FUNCTION_BLOCK "OP5_Pressure_Interlocks"
{ S7_Optimized_Access := 'TRUE' }
VERSION : 0.1
   VAR
      State {InstructionName := 'Program_Alarm'; LibVersion := '1.0'} : Program_Alarm;
      PRECOND_01 : Bool;
      PRECOND_02 : Bool;
      PRECOND_03 : Bool;
      PRECOND_04 : Bool;
      PRECOND_05 : Bool;
      PRECOND_06 : Bool;
      PRECOND_07 : Bool;
      PRECOND_08 : Bool;
      PRECOND_09 : Bool;
      PRECOND_10 : Bool;
      PRECOND_11 : Bool;
      PRECOND_12 : Bool;
      PRECOND_13 : Bool;
      PRECOND_14 : Bool;
      PRECOND_15 : Bool;
      PRECOND_16 : Bool;
      PRECOND_17 : Bool;
      PRECOND_18 : Bool;
      PRECOND_19 : Bool;
      PRECOND_20 : Bool;
      PRECOND_21 : Bool;
      PRECOND_22 : Bool;
      PRECOND_23 : Bool;
      PRECOND_24 : Bool;
      PRECOND_25 : Bool;
      PRECOND_26 : Bool;
      PRECOND_27 : Bool;
      PRECOND_28 : Bool;
      PRECOND_29 : Bool;
      PRECOND_30 : Bool;
      PRECOND_31 : Bool;
      PRECOND_32 : Bool;
      PRECOND_33 : Bool;
      PRECOND_34 : Bool;
      PRECOND_35 : Bool;
      PRECOND_36 : Bool;
      PRECOND_37 : Bool;
      PRECOND_38 : Bool;
      PRECOND_39 : Bool;
      PRECOND_40 : Bool;
      PRECOND_41 : Bool;
      PRECOND_42 : Bool;
      PRECOND_43 : Bool;
      PRECOND_44 : Bool;
      PRECOND_45 : Bool;
      PRECOND_46 : Bool;
      PRECOND_47 : Bool;
      PRECOND_48 : Bool;
      PRECOND_49 : Bool;
      PRECOND_50 : Bool;
      PH_Vent_PRECOND_01 : Bool;
      PH_Vent_PRECOND_02 : Bool;
      PH_Vent_PRECOND_03 : Bool;
      PH_Vent_PRECOND_04 : Bool;
      PH_Vent_PRECOND_05 : Bool;
      PH_Vent_PRECOND_06 : Bool;
      PH_Vent_PRECOND_07 : Bool;
      PH_Vent_PRECOND_08 : Bool;
      PH_Vent_PRECOND_09 : Bool;
      PH_Vent_PRECOND_10 : Bool;
      PH_Vent_PRECOND_11 : Bool;
      PH_Vent_PRECOND_12 : Bool;
      PH_Vent_PRECOND_13 : Bool;
      PH_Vent_PRECOND_14 : Bool;
      PH_Vent_PRECOND_15 : Bool;
      PH_Vent_PRECOND_16 : Bool;
      PH_Vent_PRECOND_17 : Bool;
      PH_Vent_PRECOND_18 : Bool;
      PH_Vent_PRECOND_19 : Bool;
      PH_Vent_PRECOND_20 : Bool;
      PH_Vent_PRECOND_21 : Bool;
      PH_Vent_PRECOND_22 : Bool;
      PH_Vent_PRECOND_23 : Bool;
      PH_Vent_PRECOND_24 : Bool;
      PH_Vent_PRECOND_25 : Bool;
      PH_Vent_PRECOND_26 : Bool;
      PH_Vent_PRECOND_27 : Bool;
      PH_Vent_PRECOND_28 : Bool;
      PH_Vent_PRECOND_29 : Bool;
      PH_Vent_PRECOND_30 : Bool;
      PH_Vent_PRECOND_31 : Bool;
      PH_Vent_PRECOND_32 : Bool;
      PH_Vent_PRECOND_33 : Bool;
      PH_Vent_PRECOND_34 : Bool;
      PH_Vent_PRECOND_35 : Bool;
      PH_Vent_PRECOND_36 : Bool;
      PH_Vent_PRECOND_37 : Bool;
      PH_Vent_PRECOND_38 : Bool;
      PH_Vent_PRECOND_39 : Bool;
      PH_Vent_PRECOND_40 : Bool;
      PH_Vent_PRECOND_41 : Bool;
      PH_Vent_PRECOND_42 : Bool;
      PH_Vent_PRECOND_43 : Bool;
      PH_Vent_PRECOND_44 : Bool;
      PH_Vent_PRECOND_45 : Bool;
      PH_Vent_PRECOND_46 : Bool;
      PH_Vent_PRECOND_47 : Bool;
      PH_Vent_PRECOND_48 : Bool;
      PH_Vent_PRECOND_49 : Bool;
      PH_Vent_PRECOND_50 : Bool;
      PH_Fill_PRECOND_01 : Bool;
      PH_Fill_PRECOND_02 : Bool;
      PH_Fill_PRECOND_03 : Bool;
      PH_Fill_PRECOND_04 : Bool;
      PH_Fill_PRECOND_05 : Bool;
      PH_Fill_PRECOND_06 : Bool;
      PH_Fill_PRECOND_07 : Bool;
      PH_Fill_PRECOND_08 : Bool;
      PH_Fill_PRECOND_09 : Bool;
      PH_Fill_PRECOND_10 : Bool;
      PH_Fill_PRECOND_11 : Bool;
      PH_Fill_PRECOND_12 : Bool;
      PH_Fill_PRECOND_13 : Bool;
      PH_Fill_PRECOND_14 : Bool;
      PH_Fill_PRECOND_15 : Bool;
      PH_Fill_PRECOND_16 : Bool;
      PH_Fill_PRECOND_17 : Bool;
      PH_Fill_PRECOND_18 : Bool;
      PH_Fill_PRECOND_19 : Bool;
      PH_Fill_PRECOND_20 : Bool;
      PH_Fill_PRECOND_21 : Bool;
      PH_Fill_PRECOND_22 : Bool;
      PH_Fill_PRECOND_23 : Bool;
      PH_Fill_PRECOND_24 : Bool;
      PH_Fill_PRECOND_25 : Bool;
      PH_Fill_PRECOND_26 : Bool;
      PH_Fill_PRECOND_27 : Bool;
      PH_Fill_PRECOND_28 : Bool;
      PH_Fill_PRECOND_29 : Bool;
      PH_Fill_PRECOND_30 : Bool;
      PH_Fill_PRECOND_31 : Bool;
      PH_Fill_PRECOND_32 : Bool;
      PH_Fill_PRECOND_33 : Bool;
      PH_Fill_PRECOND_34 : Bool;
      PH_Fill_PRECOND_35 : Bool;
      PH_Fill_PRECOND_36 : Bool;
      PH_Fill_PRECOND_37 : Bool;
      PH_Fill_PRECOND_38 : Bool;
      PH_Fill_PRECOND_39 : Bool;
      PH_Fill_PRECOND_40 : Bool;
      PH_Fill_PRECOND_41 : Bool;
      PH_Fill_PRECOND_42 : Bool;
      PH_Fill_PRECOND_43 : Bool;
      PH_Fill_PRECOND_44 : Bool;
      PH_Fill_PRECOND_45 : Bool;
      PH_Fill_PRECOND_46 : Bool;
      PH_Fill_PRECOND_47 : Bool;
      PH_Fill_PRECOND_48 : Bool;
      PH_Fill_PRECOND_49 : Bool;
      PH_Fill_PRECOND_50 : Bool;
   END_VAR

BEGIN
   REGION Function
      // here all interlocks for this operation will be defined
      // Later FALSE assignments execute every scan. Adjust them when adding calculated interlocks.
   END_REGION

   REGION General Interlocks
      #PRECOND_01 := FALSE;
      #PRECOND_02 := FALSE;
      #PRECOND_03 := FALSE;
      #PRECOND_04 := FALSE;
      #PRECOND_05 := FALSE;
      #PRECOND_06 := FALSE;
      #PRECOND_07 := FALSE;
      #PRECOND_08 := FALSE;
      #PRECOND_09 := FALSE;
      #PRECOND_10 := FALSE;
      #PRECOND_11 := FALSE;
      #PRECOND_12 := FALSE;
      #PRECOND_13 := FALSE;
      #PRECOND_14 := FALSE;
      #PRECOND_15 := FALSE;
      #PRECOND_16 := FALSE;
      #PRECOND_17 := FALSE;
      #PRECOND_18 := FALSE;
      #PRECOND_19 := FALSE;
      #PRECOND_20 := FALSE;
      #PRECOND_21 := FALSE;
      #PRECOND_22 := FALSE;
      #PRECOND_23 := FALSE;
      #PRECOND_24 := FALSE;
      #PRECOND_25 := FALSE;
      #PRECOND_26 := FALSE;
      #PRECOND_27 := FALSE;
      #PRECOND_28 := FALSE;
      #PRECOND_29 := FALSE;
      #PRECOND_30 := FALSE;
      #PRECOND_31 := FALSE;
      #PRECOND_32 := FALSE;
      #PRECOND_33 := FALSE;
      #PRECOND_34 := FALSE;
      #PRECOND_35 := FALSE;
      #PRECOND_36 := FALSE;
      #PRECOND_37 := FALSE;
      #PRECOND_38 := FALSE;
      #PRECOND_39 := FALSE;
      #PRECOND_40 := FALSE;
      #PRECOND_41 := FALSE;
      #PRECOND_42 := FALSE;
      #PRECOND_43 := FALSE;
      #PRECOND_44 := FALSE;
      #PRECOND_45 := FALSE;
      #PRECOND_46 := FALSE;
      #PRECOND_47 := FALSE;
      #PRECOND_48 := FALSE;
      #PRECOND_49 := FALSE;
      #PRECOND_50 := FALSE;
   END_REGION

   REGION PH_Vent Interlocks
      #PH_Vent_PRECOND_01 := FALSE;
      #PH_Vent_PRECOND_02 := FALSE;
      #PH_Vent_PRECOND_03 := FALSE;
      #PH_Vent_PRECOND_04 := FALSE;
      #PH_Vent_PRECOND_05 := FALSE;
      #PH_Vent_PRECOND_06 := FALSE;
      #PH_Vent_PRECOND_07 := FALSE;
      #PH_Vent_PRECOND_08 := FALSE;
      #PH_Vent_PRECOND_09 := FALSE;
      #PH_Vent_PRECOND_10 := FALSE;
      #PH_Vent_PRECOND_11 := FALSE;
      #PH_Vent_PRECOND_12 := FALSE;
      #PH_Vent_PRECOND_13 := FALSE;
      #PH_Vent_PRECOND_14 := FALSE;
      #PH_Vent_PRECOND_15 := FALSE;
      #PH_Vent_PRECOND_16 := FALSE;
      #PH_Vent_PRECOND_17 := FALSE;
      #PH_Vent_PRECOND_18 := FALSE;
      #PH_Vent_PRECOND_19 := FALSE;
      #PH_Vent_PRECOND_20 := FALSE;
      #PH_Vent_PRECOND_21 := FALSE;
      #PH_Vent_PRECOND_22 := FALSE;
      #PH_Vent_PRECOND_23 := FALSE;
      #PH_Vent_PRECOND_24 := FALSE;
      #PH_Vent_PRECOND_25 := FALSE;
      #PH_Vent_PRECOND_26 := FALSE;
      #PH_Vent_PRECOND_27 := FALSE;
      #PH_Vent_PRECOND_28 := FALSE;
      #PH_Vent_PRECOND_29 := FALSE;
      #PH_Vent_PRECOND_30 := FALSE;
      #PH_Vent_PRECOND_31 := FALSE;
      #PH_Vent_PRECOND_32 := FALSE;
      #PH_Vent_PRECOND_33 := FALSE;
      #PH_Vent_PRECOND_34 := FALSE;
      #PH_Vent_PRECOND_35 := FALSE;
      #PH_Vent_PRECOND_36 := FALSE;
      #PH_Vent_PRECOND_37 := FALSE;
      #PH_Vent_PRECOND_38 := FALSE;
      #PH_Vent_PRECOND_39 := FALSE;
      #PH_Vent_PRECOND_40 := FALSE;
      #PH_Vent_PRECOND_41 := FALSE;
      #PH_Vent_PRECOND_42 := FALSE;
      #PH_Vent_PRECOND_43 := FALSE;
      #PH_Vent_PRECOND_44 := FALSE;
      #PH_Vent_PRECOND_45 := FALSE;
      #PH_Vent_PRECOND_46 := FALSE;
      #PH_Vent_PRECOND_47 := FALSE;
      #PH_Vent_PRECOND_48 := FALSE;
      #PH_Vent_PRECOND_49 := FALSE;
      #PH_Vent_PRECOND_50 := FALSE;
   END_REGION

   REGION PH_Fill Interlocks
      #PH_Fill_PRECOND_01 := FALSE;
      #PH_Fill_PRECOND_02 := FALSE;
      #PH_Fill_PRECOND_03 := FALSE;
      #PH_Fill_PRECOND_04 := FALSE;
      #PH_Fill_PRECOND_05 := FALSE;
      #PH_Fill_PRECOND_06 := FALSE;
      #PH_Fill_PRECOND_07 := FALSE;
      #PH_Fill_PRECOND_08 := FALSE;
      #PH_Fill_PRECOND_09 := FALSE;
      #PH_Fill_PRECOND_10 := FALSE;
      #PH_Fill_PRECOND_11 := FALSE;
      #PH_Fill_PRECOND_12 := FALSE;
      #PH_Fill_PRECOND_13 := FALSE;
      #PH_Fill_PRECOND_14 := FALSE;
      #PH_Fill_PRECOND_15 := FALSE;
      #PH_Fill_PRECOND_16 := FALSE;
      #PH_Fill_PRECOND_17 := FALSE;
      #PH_Fill_PRECOND_18 := FALSE;
      #PH_Fill_PRECOND_19 := FALSE;
      #PH_Fill_PRECOND_20 := FALSE;
      #PH_Fill_PRECOND_21 := FALSE;
      #PH_Fill_PRECOND_22 := FALSE;
      #PH_Fill_PRECOND_23 := FALSE;
      #PH_Fill_PRECOND_24 := FALSE;
      #PH_Fill_PRECOND_25 := FALSE;
      #PH_Fill_PRECOND_26 := FALSE;
      #PH_Fill_PRECOND_27 := FALSE;
      #PH_Fill_PRECOND_28 := FALSE;
      #PH_Fill_PRECOND_29 := FALSE;
      #PH_Fill_PRECOND_30 := FALSE;
      #PH_Fill_PRECOND_31 := FALSE;
      #PH_Fill_PRECOND_32 := FALSE;
      #PH_Fill_PRECOND_33 := FALSE;
      #PH_Fill_PRECOND_34 := FALSE;
      #PH_Fill_PRECOND_35 := FALSE;
      #PH_Fill_PRECOND_36 := FALSE;
      #PH_Fill_PRECOND_37 := FALSE;
      #PH_Fill_PRECOND_38 := FALSE;
      #PH_Fill_PRECOND_39 := FALSE;
      #PH_Fill_PRECOND_40 := FALSE;
      #PH_Fill_PRECOND_41 := FALSE;
      #PH_Fill_PRECOND_42 := FALSE;
      #PH_Fill_PRECOND_43 := FALSE;
      #PH_Fill_PRECOND_44 := FALSE;
      #PH_Fill_PRECOND_45 := FALSE;
      #PH_Fill_PRECOND_46 := FALSE;
      #PH_Fill_PRECOND_47 := FALSE;
      #PH_Fill_PRECOND_48 := FALSE;
      #PH_Fill_PRECOND_49 := FALSE;
      #PH_Fill_PRECOND_50 := FALSE;
   END_REGION
END_FUNCTION_BLOCK
